Yaskawa INFORM job: 1-DEFRO-5.JBI

/JOB
//NAME 1-DEFRO-5
//POS
///NPOS 9,9,9,0,0,0
///TOOL 0
///POSTYPE PULSE
///PULSE
C00000=-283,-101162,-84213,3710,-80188,-1936
C00001=-275,-97864,-82985,3720,-79251,-1967
C00002=-100003,31603,4033,-7680,-72698,-47529
C00003=-94834,78089,9543,-9078,-51926,-47788
C00004=-83555,68320,-11474,26050,-31610,-59171
C00005=-83555,68320,-11474,26050,-31610,-59171
C00006=-102318,64841,-853,-9216,-53032,-45265
C00007=-275,-97864,-82985,3720,-79251,-1967
C00008=-283,-101162,-84213,3710,-80188,-1936
BC00000=570125
BC00001=808681
BC00002=808681
BC00003=808681
BC00004=808680
BC00005=808680
BC00006=808681
BC00007=808681
BC00008=570125
EC00000=1,-94526
EC00001=1,-94526
EC00002=1,-94526
EC00003=1,-94526
EC00004=-2638,-94527
EC00005=-2638,-726117
EC00006=-73,-613687
EC00007=1,-94526
EC00008=1,-94526
//INST
///DATE 2025/01/13 12:40
///ATTR SC,RW
///GROUP1 RB1,BS1
///GROUP2 ST3
NOP
MOVJ C00000 BC00000 VJ=40.00 DEC=20  +MOVJ EC00000 VJ=40.00
MOVJ C00001 BC00001 VJ=40.00 DEC=20  +MOVJ EC00001 VJ=40.00
MOVJ C00002 BC00002 VJ=40.00 DEC=20  +MOVJ EC00002 VJ=40.00
MOVJ C00003 BC00003 VJ=40.00 DEC=20  +MOVJ EC00003 VJ=40.00
MOVJ C00004 BC00004 VJ=40.00 DEC=20  +MOVJ EC00004 VJ=40.00
MACRO1 MJ#(0) ARGF4
ARCON
MOVJ C00005 BC00005 VJ=0.78 DEC=20  +MOVJ EC00005 VJ=20.00
ARCOF
MOVJ C00006 BC00006 VJ=40.00 DEC=20  +MOVJ EC00006 VJ=40.00
MOVJ C00007 BC00007 VJ=40.00 DEC=20  +MOVJ EC00007 VJ=40.00
MOVJ C00008 BC00008 VJ=40.00 DEC=20  +MOVJ EC00008 VJ=40.00
END
